Fanuc KAREL source: kt00473.KL

-- PROVISIONAL review KL for V770-1; original PC SHA256 1281a5dc7c13b85318edbaa82ae8e9b725934e4130e9f272491d120ce95a4ab2
-- Incomplete behavior may be omitted. Consult companion uncertainty JSON. Do not deploy.
PROGRAM KT00473
%NOLOCKGROUP
VAR
  OUT : BOOLEAN
-- UNRESOLVED_DECL P1 type=000101
-- UNRESOLVED_DECL P2 type=000101
BEGIN
  -- UNRESOLVED_PC offsets 5-28; opcodes 49,49,AC,23
  -- UNRESOLVED_PC offsets 33-37; opcodes 7F
END KT00473
